// TIA Portal V19 export
TYPE "EM01_Input"
   STRUCT
      Cmds { S7_SetPoint := 'True'} : "EM_Input";
      CtrlMode : Int;   // 0=Off, 1=Calentamiento por temperatura, 2=Local (concentraciÃ³n), 3=External (SeedMaster), 4=Limpieza/caldeo por tiempo, 5=Lavado por tiempo
      TempSP : Real;
      TempFilter : Time := T#3S;   // Tiempo que PV >= SP debe mantenerse para completar
      TimeSP : Time;
      Timeout : Time;   // Tiempo mÃ¡ximo para alcanzar la temperatura
      ValveTime : Time := T#10S;   // Tiempo mÃ¡ximo de confirmaciÃ³n de apertura/cierre de la vÃ¡lvula
      ConcentrationSP : Real;   // SP de concentraciÃ³n/Brix (0..100); objetivo en modos 2 y 3
      ConcStableBand : Real := 1.0;   // Banda de estabilizaciÃ³n de concentraciÃ³n (modos 2 y 3)
      ConcStableTime : Time := T#30S;   // Tiempo dentro de banda para declarar COMPLETED (modos 2 y 3)
      ConcSMMV : Real;   // MV del SeedMaster en % (0..100), modo 3
      HoldPosition : Real;   // PosiciÃ³n fija del PID en Hold/Held, % (0..100), modos 2 y 3
      MinLevelPermit : Bool;   // Nivel de tacho suficiente para cubrir la calandria
      DischargeInterlock : Bool;   // TRUE durante la descarga: calandria forzada a 0 %
   END_STRUCT;
END_TYPE
